Staubli VAL3: onSave.pgx

public program onSave(bool& x_bToSave)
begin
  if x_bToSave
    rs:bIsSaving=true
    trajTemp:libSave()
    x_bToSave=false
    rs:bIsSaving=false
    delay(0.5)
    popUpMsg("trajectory数据已保存")
  endIf
end
